% RSLogix 500 project PROGRAM 3.RSS, saved by version 8.30.00.16 %
PROJECT "UNTITLED"    % processor: Bul.1763 MicroLogix 1100 Series B %

PROGRAM FILES
  LAD 2 "MAIN"  2 rungs
  LAD 3 "BARCODE"  6 rungs
  LAD 4 "INVENTORY"  8 rungs

DATA FILES
  O0 OUTPUT  4 elements
  I1 INPUT  6 elements
  S2 STATUS  66 elements
  B3 BINARY  1 elements
  T4 TIMER  1 elements
  C5 COUNTER  1 elements
  R6 CONTROL  1 elements
  N7 INTEGER  6 elements
  F8 FLOAT  1 elements
  ST9 STRING  4 elements

LADDER 2 "MAIN"
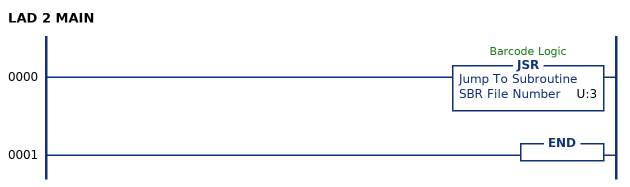
% Rung: 0 %
SOR JSR U:3 EOR
%   U:3  "Barcode Logic" %
% Rung: 1 %
SOR END EOR

LADDER 3 "BARCODE"
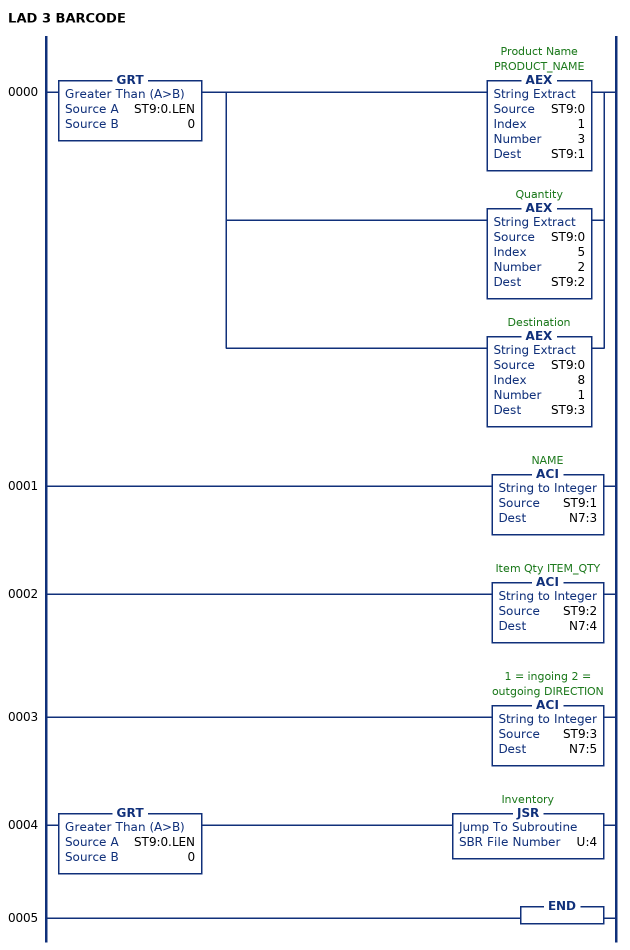
% Rung: 0 %
SOR GRT ST9:0.LEN 0 BST AEX ST9:0 1 3 ST9:1 NXB AEX ST9:0 5 2 ST9:2 NXB AEX ST9:0 8 1 ST9:3 BND EOR
%   ST9:0  ST9  "Barcode Scanner" %
%   ST9:1  PRODUCT_NAME  "Product Name" %
%   ST9:2  "Quantity" %
%   ST9:3  "Destination" %
% Rung: 1 %
SOR ACI ST9:1 N7:3 EOR
%   ST9:1  PRODUCT_NAME  "Product Name" %
%   N7:3  NAME %
% Rung: 2 %
SOR ACI ST9:2 N7:4 EOR
%   ST9:2  "Quantity" %
%   N7:4  ITEM_QTY  "Item Qty" %
% Rung: 3 %
SOR ACI ST9:3 N7:5 EOR
%   ST9:3  "Destination" %
%   N7:5  DIRECTION  "1 = ingoing 2 = outgoing" %
% Rung: 4 %
SOR GRT ST9:0.LEN 0 JSR U:4 EOR
%   U:4  "Inventory" %
% Rung: 5 %
SOR END EOR

LADDER 4 "INVENTORY"
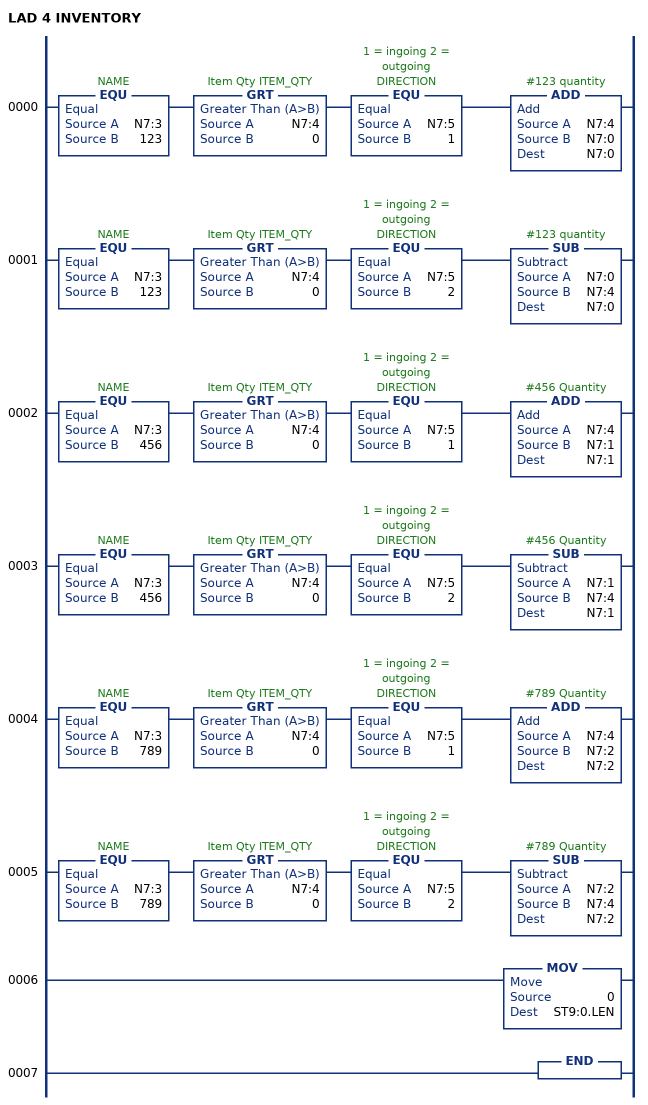
% Rung: 0 %
SOR EQU N7:3 123 GRT N7:4 0 EQU N7:5 1 ADD N7:4 N7:0 N7:0 EOR
%   N7:3  NAME %
%   N7:4  ITEM_QTY  "Item Qty" %
%   N7:5  DIRECTION  "1 = ingoing 2 = outgoing" %
%   N7:0  "#123 quantity" %
% Rung: 1 %
SOR EQU N7:3 123 GRT N7:4 0 EQU N7:5 2 SUB N7:0 N7:4 N7:0 EOR
%   N7:3  NAME %
%   N7:4  ITEM_QTY  "Item Qty" %
%   N7:5  DIRECTION  "1 = ingoing 2 = outgoing" %
%   N7:0  "#123 quantity" %
% Rung: 2 %
SOR EQU N7:3 456 GRT N7:4 0 EQU N7:5 1 ADD N7:4 N7:1 N7:1 EOR
%   N7:3  NAME %
%   N7:4  ITEM_QTY  "Item Qty" %
%   N7:5  DIRECTION  "1 = ingoing 2 = outgoing" %
%   N7:1  "#456 Quantity" %
% Rung: 3 %
SOR EQU N7:3 456 GRT N7:4 0 EQU N7:5 2 SUB N7:1 N7:4 N7:1 EOR
%   N7:3  NAME %
%   N7:4  ITEM_QTY  "Item Qty" %
%   N7:5  DIRECTION  "1 = ingoing 2 = outgoing" %
%   N7:1  "#456 Quantity" %
% Rung: 4 %
SOR EQU N7:3 789 GRT N7:4 0 EQU N7:5 1 ADD N7:4 N7:2 N7:2 EOR
%   N7:3  NAME %
%   N7:4  ITEM_QTY  "Item Qty" %
%   N7:5  DIRECTION  "1 = ingoing 2 = outgoing" %
%   N7:2  "#789 Quantity" %
% Rung: 5 %
SOR EQU N7:3 789 GRT N7:4 0 EQU N7:5 2 SUB N7:2 N7:4 N7:2 EOR
%   N7:3  NAME %
%   N7:4  ITEM_QTY  "Item Qty" %
%   N7:5  DIRECTION  "1 = ingoing 2 = outgoing" %
%   N7:2  "#789 Quantity" %
% Rung: 6 %
SOR MOV 0 ST9:0.LEN EOR
% Rung: 7 %
SOR END EOR

OTHER DOCUMENTED ADDRESSES
  B3:0/0  "ONS"
  B3:0/1  "ONS"

DATA TABLE (non-zero values as saved)
DATA N7
% N7:0 % 0 0 70 789 80 1
DATA ST9
% ST9:1 % "789"
% ST9:2 % "80"
% ST9:3 % "1"
